Fanuc KAREL source: KB00101.KL

PROGRAM KB00101
%NOLOCKGROUP
%ENVIRONMENT UIF
VAR
  P1: INTEGER
  P2: STRING[80]
  P3: INTEGER
  P4: INTEGER
  P5: INTEGER
  P6: INTEGER
  P7: INTEGER
  P8: INTEGER
  P9: ARRAY[4] OF STRING[80]
  P10: INTEGER
BEGIN
  P1 = 1
  P2 = 'A'
  P3 = 1
  P4 = 1
  P5 = 1
  P6 = 1
  P7 = 1
  P8 = 1
  P10 = 1
  INI_DYN_DISE(P1, P2, P3, P4, P5, P6, P7, P8, P9, P10)
END KB00101
